Fanuc KAREL source: KA00188.KL

PROGRAM KA00188
%NOLOCKGROUP
VAR
  SRC: ARRAY[4] OF BYTE
  DST: ARRAY[4] OF XYZWPR
BEGIN
  DST = SRC
END KA00188
